(* IEC 61131-3 sources: kns-port-domestic/upstream/kns-pump-station/src/POUs/Station/FB_ControlSelector, 2 files *)

(* ---- FB_ControlSelector.decl.st ---- *)
// Назначение: действующее управление насосами (04 §4). В «Автомате» по старшинству: PowerLost >
//             Restart > DryRunStop > Float > Emergency > LevelPid (выбран и готов) > Stepped; в
//             «Ручном» — Manual. xStepFallback — условие тревоги KNS1.STEP (выбран ПИД, ПИД не
//             готов); xChanged — импульс смены управления (вход без рывка в PRG_Station).
// Автор:      kr0nsch
// Версия:     0.1.0
// Документ:   docs/DESIGN.md, раздел 6.2; docs/04_algorithms.md, раздел 4
FUNCTION_BLOCK FB_ControlSelector
VAR_INPUT
    eMode      : E_StationMode;
    eMethod    : E_ControlMethod;
    xPowerLost : BOOL;              // FB_PowerRestore
    xRestart   : BOOL;
    xDryRun    : BOOL;              // FB_Protections
    xFloatMode : BOOL;
    xEmergency : BOOL;
    xPidReady  : BOOL;              // FB_LevelControlPid
END_VAR
VAR_OUTPUT
    eControlAct   : E_ControlAct;
    xStepFallback : BOOL;           // Auto, выбран ПИД, ПИД не готов (условие KNS1.STEP)
    xChanged      : BOOL;           // eControlAct сменилось в этом вызове
END_VAR
VAR
    eActPrev : E_ControlAct;        // управление прошлого вызова (первый вызов — Manual)
END_VAR

(* ---- FB_ControlSelector.impl.st ---- *)
// Режим вне перечисления (мусор) — как «Ручной», способ вне перечисления — как «Ступенчатое»
// (E_StationMode, E_ControlMethod: безопасный вариант)
IF eMode <> E_StationMode.Auto THEN
    eControlAct := E_ControlAct.Manual;
ELSIF xPowerLost THEN
    eControlAct := E_ControlAct.PowerLost;
ELSIF xRestart THEN
    eControlAct := E_ControlAct.Restart;
ELSIF xDryRun THEN
    eControlAct := E_ControlAct.DryRunStop;
ELSIF xFloatMode THEN
    eControlAct := E_ControlAct.Float;
ELSIF xEmergency THEN
    eControlAct := E_ControlAct.Emergency;
ELSIF eMethod = E_ControlMethod.LevelPid AND xPidReady THEN
    eControlAct := E_ControlAct.LevelPid;
ELSE
    eControlAct := E_ControlAct.Stepped;
END_IF

// Условие KNS1.STEP не зависит от старших состояний: их подавление задаёт PRG_Station (04 §15)
xStepFallback := eMode = E_StationMode.Auto AND eMethod = E_ControlMethod.LevelPid AND NOT xPidReady;

xChanged := eControlAct <> eActPrev;
eActPrev := eControlAct;
